(* IEC 61131-3 sources: RootPLC/crates/rootplc-stdlib/libs/Tc3_EventLogger/1.0.0, 1 file *)

(* ---- Tc3_EventLogger.st ---- *)
(* Tc3_EventLogger compatibility library for RootPLC (see library.toml).

   Written from the public library manual (TE1000 PLC Library:
   Tc3_EventLogger, version 1.6.2). RootPLC has no TwinCAT EventLogger
   service, so the blocks that talk to it are declared but not implemented
   (library.toml declare_only): calls type-check and give warning RP0120, and
   running one stops with UNSUPPORTED. FB_TcSourceInfo holds data only and is
   implemented, except ResetToDefault (it needs the instance's symbol name).

   Differences from the manual, all because the manual does not publish the
   definition:
   - interfaces used only as parameter or property types (filter
     expressions, remote logger, listener context, export settings) are
     declared without members;
   - FB_TcEventFilter has only the members the manual lists;
     FB_TcClearLoggedEventsSettings lacks SetLimit / SetSorting; the remote
     logger blocks and the ADS error conversions (E_AdsErr,
     E_HRESULTAdsErr) are left out;
   - sName of the source information is STRING(255): the manual's
     STRING(ParameterList.cSourceNameSize - 1) with the default size 256.
   TC_EVENTS is generated by TwinCAT from the project's event classes and
   is not part of this library. *)

{attribute 'qualified_only'}
TYPE TcEventSeverity : (
    Verbose  := 0,
    Info     := 1,
    Warning  := 2,
    Error    := 3,
    Critical := 4);
END_TYPE

{attribute 'qualified_only'}
TYPE TcEventConfirmationState : (
    NotSupported := 0,
    NotRequired  := 1,
    WaitForConfirmation := 2,
    Confirmed := 3,
    Reset     := 4);
END_TYPE

TYPE TcEventEntry :
STRUCT
    uuidEventClass : GUID;
    nEventId       : UDINT;
    eSeverity      : TcEventSeverity;
END_STRUCT
END_TYPE

VAR_GLOBAL CONSTANT
    EMPTY_EVENT_CLASS : GUID := (Data1 := 16#0, Data2 := 16#0, Data3 := 16#0, Data4 := [16#0, 16#0, 16#0, 16#0, 16#0, 16#0, 16#0, 16#0]);
    EMPTY_EVENT_ID    : UDINT := 16#0;
    EMPTY_SEVERITY    : TcEventSeverity := TcEventSeverity#Verbose;
    SUCCESS_EVENT     : TcEventEntry := (uuidEventClass := EMPTY_EVENT_CLASS, nEventId := EMPTY_EVENT_ID, eSeverity := EMPTY_SEVERITY);
    stLibVersion_Tc3_EventLogger : ST_LibVersion;
END_VAR

NAMESPACE GVL
VAR_GLOBAL
    nLangId_OnlineMonitoring : DINT := 1033;
END_VAR
END_NAMESPACE

NAMESPACE ParameterList
VAR_GLOBAL CONSTANT
    cSourceNameSize : UDINT(81..10000) := 256;
END_VAR
END_NAMESPACE

(* interfaces the manual names without publishing their members *)
INTERFACE I_TcRemoteEventLogger
END_INTERFACE
INTERFACE I_TcListenerContext
END_INTERFACE
INTERFACE I_TcEventFilterBase
END_INTERFACE
INTERFACE I_TcEventFilter EXTENDS I_TcEventFilterBase
END_INTERFACE
INTERFACE I_TcExpressionBase
END_INTERFACE
INTERFACE I_TcBinaryExpression
END_INTERFACE
INTERFACE I_TcLogicalExpression
END_INTERFACE
INTERFACE I_TcAlarmFilterExpression
END_INTERFACE
INTERFACE I_TcEtherCATDeviceExpression
END_INTERFACE
INTERFACE I_TcGuidCompare
END_INTERFACE
INTERFACE I_TcUDIntCompare
END_INTERFACE
INTERFACE I_TcULIntCompare
END_INTERFACE
INTERFACE I_TcJsonAttributeExpression
END_INTERFACE
INTERFACE I_TcSeverityCompare
END_INTERFACE
INTERFACE I_TcSourceInfoExpression
END_INTERFACE
INTERFACE I_TcClearLoggedEventsSettings
END_INTERFACE
INTERFACE I_TcEventExportSettings
END_INTERFACE
INTERFACE ITcEventFilterConfig
END_INTERFACE

INTERFACE I_TcSourceInfo
METHOD EqualsTo : BOOL
VAR_INPUT
    ipOther : I_TcSourceInfo;
END_VAR
END_METHOD
PROPERTY guid : GUID
GET
END_GET
END_PROPERTY
PROPERTY nId : UDINT
GET
END_GET
END_PROPERTY
PROPERTY sName : STRING(255)
GET
END_GET
END_PROPERTY
END_INTERFACE

INTERFACE I_TcArguments
METHOD AddBlob : I_TcArguments
VAR_INPUT
    pData  : PVOID;
    cbData : UINT;
END_VAR
END_METHOD
METHOD AddBool : I_TcArguments
VAR_INPUT
    value : BOOL;
END_VAR
END_METHOD
METHOD AddByte : I_TcArguments
VAR_INPUT
    value : BYTE;
END_VAR
END_METHOD
METHOD AddDINT : I_TcArguments
VAR_INPUT
    value : DINT;
END_VAR
END_METHOD
METHOD AddDWord : I_TcArguments
VAR_INPUT
    value : DWORD;
END_VAR
END_METHOD
METHOD AddEventReferenceId : I_TcArguments
VAR_INPUT
    nEventId : UDINT;
END_VAR
END_METHOD
METHOD AddEventReferenceIdGuid : I_TcArguments
VAR_INPUT
    nEventId   : UDINT;
    EventClass : GUID;
END_VAR
END_METHOD
METHOD AddINT : I_TcArguments
VAR_INPUT
    value : INT;
END_VAR
END_METHOD
METHOD AddLInt : I_TcArguments
VAR_INPUT
    value : LINT;
END_VAR
END_METHOD
METHOD AddLReal : I_TcArguments
VAR_INPUT
    value : LREAL;
END_VAR
END_METHOD
METHOD AddReal : I_TcArguments
VAR_INPUT
    value : REAL;
END_VAR
END_METHOD
METHOD AddSInt : I_TcArguments
VAR_INPUT
    value : SInt;
END_VAR
END_METHOD
METHOD AddString : I_TcArguments
VAR_IN_OUT CONSTANT
    value : STRING;
END_VAR
END_METHOD
METHOD AddUDInt : I_TcArguments
VAR_INPUT
    value : UDINT;
END_VAR
END_METHOD
METHOD AddUInt : I_TcArguments
VAR_INPUT
    value : UINT;
END_VAR
END_METHOD
METHOD AddULInt : I_TcArguments
VAR_INPUT
    value : ULINT;
END_VAR
END_METHOD
METHOD AddUSInt : I_TcArguments
VAR_INPUT
    value : USINT;
END_VAR
END_METHOD
METHOD AddWord : I_TcArguments
VAR_INPUT
    value : WORD;
END_VAR
END_METHOD
METHOD AddWString : I_TcArguments
VAR_IN_OUT CONSTANT
    value : WSTRING;
END_VAR
END_METHOD
METHOD Clear : I_TcArguments
END_METHOD
PROPERTY nCount : UDINT
GET
END_GET
END_PROPERTY
END_INTERFACE

INTERFACE I_TcEventBase
METHOD EqualsTo : BOOL
VAR_INPUT
    ipOther : I_TcEventBase;
END_VAR
END_METHOD
METHOD EqualsToEventClass : BOOL
VAR_INPUT
    OtherEventClass : GUID;
END_VAR
END_METHOD
METHOD EqualsToEventEntry : BOOL
VAR_INPUT
    OtherEventClass : GUID;
    nOtherEventID   : UDINT;
    eOtherSeverity  : TcEventSeverity;
END_VAR
END_METHOD
METHOD EqualsToEventEntryEx : BOOL
VAR_INPUT
    stOther : TcEventEntry;
END_VAR
END_METHOD
METHOD GetJsonAttribute : HRESULT
VAR_INPUT
    sJsonAttribute : REFERENCE TO STRING;
    nJsonAttribute : UDINT;
END_VAR
END_METHOD
METHOD RequestEventClassName : BOOL
VAR_INPUT
    nLangId     : DINT;
    sResult     : REFERENCE TO STRING;
    nResultSize : UDINT;
END_VAR
VAR_OUTPUT
    bError      : BOOL;
    hrErrorCode : HRESULT;
END_VAR
END_METHOD
METHOD RequestEventText : BOOL
VAR_INPUT
    nLangId     : DINT;
    sResult     : REFERENCE TO STRING;
    nResultSize : UDINT;
END_VAR
VAR_OUTPUT
    bError      : BOOL;
    hrErrorCode : HRESULT;
END_VAR
END_METHOD
PROPERTY eSeverity : TcEventSeverity
GET
END_GET
END_PROPERTY
PROPERTY EventClass : GUID
GET
END_GET
END_PROPERTY
PROPERTY ipSourceInfo : I_TcSourceInfo
GET
END_GET
END_PROPERTY
PROPERTY nEventId : UDINT
GET
END_GET
END_PROPERTY
PROPERTY stEventEntry : TcEventEntry
GET
END_GET
END_PROPERTY
END_INTERFACE

INTERFACE I_TcMessage EXTENDS I_TcEventBase
METHOD Send : HRESULT
VAR_INPUT
    nTimeStamp: ULINT;
END_VAR
END_METHOD
END_INTERFACE

INTERFACE I_Listener2
METHOD OnAlarmCleared : HRESULT
VAR_INPUT
    fbEvent : REFERENCE TO FB_TcEvent;
END_VAR
END_METHOD
METHOD OnAlarmConfirmed : HRESULT
VAR_INPUT
    fbEvent : REFERENCE TO FB_TcEvent;
END_VAR
END_METHOD
METHOD OnAlarmDisposed : HRESULT
VAR_INPUT
    fbEvent : REFERENCE TO FB_TcEvent;
END_VAR
END_METHOD
METHOD OnAlarmRaised : HRESULT
VAR_INPUT
    fbEvent : REFERENCE TO FB_TcEvent;
END_VAR
END_METHOD
METHOD OnMessageSent : HRESULT
VAR_INPUT
    fbEvent : REFERENCE TO FB_TcEvent;
END_VAR
END_METHOD
END_INTERFACE

FUNCTION_BLOCK FB_AsyncStrResult
METHOD GetString : BOOL
VAR_INPUT
    sResult : REFERENCE TO STRING;
    nResult : UDINT;
END_VAR
END_METHOD
PROPERTY bBusy : BOOL
GET
END_GET
END_PROPERTY
PROPERTY bError : BOOL
GET
END_GET
END_PROPERTY
PROPERTY hrErrorCode : HRESULT
GET
END_GET
END_PROPERTY
END_FUNCTION_BLOCK

FUNCTION_BLOCK FB_TcCauseRemedy
METHOD GetCause : BOOL
VAR_INPUT
    sResult     : REFERENCE TO STRING;
    nResult     : UDINT; (* buffer size in bytes *)
END_VAR
END_METHOD
METHOD GetId : BOOL
VAR_INPUT
    sResult  : REFERENCE TO STRING;
    nResult  : UDINT; (* buffer size in bytes *)
END_VAR
END_METHOD
METHOD GetRemedy : BOOL
VAR_INPUT
    sResult      : REFERENCE TO STRING;
    nResult      : UDINT; (* buffer size in bytes *)
END_VAR
END_METHOD
METHOD Release : HRESULT
END_METHOD
END_FUNCTION_BLOCK

FUNCTION_BLOCK FB_TcDetail
METHOD Release : HRESULT
END_METHOD
METHOD GetComment : BOOL
VAR_INPUT
    sResult       : REFERENCE TO STRING;
    nResult       : UDINT; (* buffer size in bytes *)
END_VAR
END_METHOD
METHOD GetName : BOOL
VAR_INPUT
    sResult    : REFERENCE TO STRING;
    nResult    : UDINT; (* buffer size in bytes *)
END_VAR
END_METHOD
METHOD GetText : BOOL
VAR_INPUT
    sResult    : REFERENCE TO STRING;
    nResult    : UDINT; (* buffer size in bytes *)
END_VAR
END_METHOD
END_FUNCTION_BLOCK

FUNCTION_BLOCK FB_RequestCauseRemedy
METHOD Clear
END_METHOD
METHOD Get        : HRESULT
VAR_INPUT
    nIndex        : UDINT;
    fbCauseRemedy : REFERENCE TO FB_TcCauseRemedy;
END_VAR
END_METHOD
METHOD Request : HRESULT
VAR_INPUT
    eventClass : GUID;
    nEventId   : UDINT;
    nLangId    : DINT; (* English(US)=1033 ; German(Germay)=1031 *)
END_VAR
END_METHOD
METHOD RequestRemote : HRESULT
VAR_INPUT
    ipRemoteLogger   : I_TcRemoteEventLogger;
    eventClass       : GUID;
    nEventId         : UDINT;
    nLangId          : DINT; (* English(US)=1033 ; German(Germay)=1031 *)
END_VAR
END_METHOD
PROPERTY bBusy : BOOL
GET
END_GET
END_PROPERTY
PROPERTY bError : BOOL
GET
END_GET
END_PROPERTY
PROPERTY hrErrorCode : HRESULT
GET
END_GET
END_PROPERTY
PROPERTY nCount : UDINT
GET
END_GET
END_PROPERTY
END_FUNCTION_BLOCK

FUNCTION_BLOCK FB_RequestEventClassDetails
METHOD Clear
END_METHOD
METHOD Get   : HRESULT
VAR_INPUT
    nIndex   : UDINT;
    fbDetail : REFERENCE TO FB_TcDetail;
END_VAR
END_METHOD
METHOD Request : HRESULT
VAR_INPUT
    eventClass : GUID;
    nLangId    : DINT; (* English(US)=1033 ; German(Germay)=1031 *)
END_VAR
END_METHOD
METHOD RequestRemote : HRESULT
VAR_INPUT
    ipRemoteLogger   : I_TcRemoteEventLogger;
    eventClass       : GUID;
    nLangId          : DINT; (* English(US)=1033 ; German(Germay)=1031 *)
END_VAR
END_METHOD
PROPERTY bBusy : BOOL
GET
END_GET
END_PROPERTY
PROPERTY bError : BOOL
GET
END_GET
END_PROPERTY
PROPERTY hrErrorCode : HRESULT
GET
END_GET
END_PROPERTY
PROPERTY nCount : UDINT
GET
END_GET
END_PROPERTY
END_FUNCTION_BLOCK

FUNCTION_BLOCK FB_RequestEventClassName
METHOD Clear
END_METHOD
METHOD GetString : BOOL
VAR_INPUT
    sResult : REFERENCE TO STRING;
    nResult : UDINT;
END_VAR
END_METHOD
METHOD Request : HRESULT
VAR_INPUT
    eventClass : GUID;
    nLangId    : DINT;
END_VAR
END_METHOD
METHOD RequestRemote : HRESULT
VAR_INPUT
    ipRemoteLogger   : I_TcRemoteEventLogger;
    eventClass       : GUID;
    nLangId          : DINT; (* English(US)=1033 ; German(Germay)=1031 *)
END_VAR
END_METHOD
PROPERTY bBusy : BOOL
GET
END_GET
END_PROPERTY
PROPERTY bError : BOOL
GET
END_GET
END_PROPERTY
PROPERTY hrErrorCode : HRESULT
GET
END_GET
END_PROPERTY
END_FUNCTION_BLOCK

FUNCTION_BLOCK FB_RequestEventDetails
METHOD Clear
END_METHOD
METHOD Get   : HRESULT
VAR_INPUT
    nIndex   : UDINT;
    fbDetail : REFERENCE TO FB_TcDetail;
END_VAR
END_METHOD
METHOD Request : HRESULT
VAR_INPUT
    eventClass : GUID;
    nEventId   : UDINT;
    nLangId    : DINT; (* English(US)=1033 ; German(Germay)=1031 *)
END_VAR
END_METHOD
METHOD RequestRemote : HRESULT
VAR_INPUT
    ipRemoteLogger   : I_TcRemoteEventLogger;
    eventClass       : GUID;
    nEventId         : UDINT;
    nLangId          : DINT; (* English(US)=1033 ; German(Germay)=1031 *)
END_VAR
END_METHOD
PROPERTY bBusy : BOOL
GET
END_GET
END_PROPERTY
PROPERTY bError : BOOL
GET
END_GET
END_PROPERTY
PROPERTY hrErrorCode : HRESULT
GET
END_GET
END_PROPERTY
PROPERTY nCount : UDINT
GET
END_GET
END_PROPERTY
END_FUNCTION_BLOCK

FUNCTION_BLOCK FB_RequestEventText
METHOD GetString : BOOL
VAR_INPUT
    sResult : REFERENCE TO STRING;
    nResult : UDINT;
END_VAR
END_METHOD
METHOD Request : BOOL
VAR_INPUT
    eventClass : GUID;
    nEventId   : UDINT;
    nLangId    : DINT;
    ipArgs     : I_TcArguments;
END_VAR
END_METHOD
METHOD RequestRemote : HRESULT
VAR_INPUT
    ipRemoteLogger   : I_TcRemoteEventLogger;
    eventClass       : GUID;
    nEventId         : UDINT;
    nLangId          : DINT;
    ipArgs           : I_TcArguments;
END_VAR
END_METHOD
METHOD Clear
END_METHOD
PROPERTY bBusy : BOOL
GET
END_GET
END_PROPERTY
PROPERTY bError : BOOL
GET
END_GET
END_PROPERTY
PROPERTY hrErrorCode : HRESULT
GET
END_GET
END_PROPERTY
END_FUNCTION_BLOCK

FUNCTION_BLOCK FB_RequestTranslation
METHOD GetString : BOOL
VAR_INPUT
    sResult : REFERENCE TO STRING;
    nResult : UDINT;
END_VAR
END_METHOD
METHOD Request : BOOL
VAR_INPUT
    eventClass : GUID;
END_VAR
VAR_IN_OUT CONSTANT
    text       : STRING;
END_VAR
VAR_INPUT
    nLangId    : DINT;
    ipArgs     : I_TcArguments;
END_VAR
END_METHOD
METHOD RequestRemote : HRESULT
VAR_INPUT
    ipRemoteLogger   : I_TcRemoteEventLogger;
    eventClass       : GUID;
END_VAR
VAR_IN_OUT CONSTANT
    text             : STRING;
END_VAR
VAR_INPUT
    nLangId          : DINT;
    ipArgs           : I_TcArguments;
END_VAR
END_METHOD
METHOD Clear
END_METHOD
PROPERTY bBusy : BOOL
GET
END_GET
END_PROPERTY
PROPERTY bError : BOOL
GET
END_GET
END_PROPERTY
PROPERTY hrErrorCode : HRESULT
GET
END_GET
END_PROPERTY
END_FUNCTION_BLOCK

FUNCTION_BLOCK FB_TcEventBase
METHOD EqualsTo : BOOL
VAR_INPUT
    ipOther : I_TcEventBase;
END_VAR
END_METHOD
METHOD EqualsToEventClass : BOOL
VAR_INPUT
    OtherEventClass : GUID;
END_VAR
END_METHOD
METHOD EqualsToEventEntry : BOOL
VAR_INPUT
    OtherEventClass : GUID;
    nOtherEventID   : UDINT;
    eOtherSeverity  : TcEventSeverity;
END_VAR
END_METHOD
METHOD EqualsToEventEntryEx : BOOL
VAR_INPUT
    stOther : TcEventEntry;
END_VAR
END_METHOD
METHOD GetJsonAttribute : HRESULT
VAR_INPUT
    sJsonAttribute : REFERENCE TO STRING;
    nJsonAttribute : UDINT;
END_VAR
END_METHOD
METHOD Release : HRESULT
END_METHOD
METHOD RequestEventClassName : BOOL
VAR_INPUT
    nLangId     : DINT;
    sResult     : REFERENCE TO STRING;
    nResultSize : UDINT;
END_VAR
VAR_OUTPUT
    bError      : BOOL;
    hrErrorCode : HRESULT;
END_VAR
END_METHOD
METHOD RequestEventText : BOOL
VAR_INPUT
    nLangId     : DINT;
    sResult     : REFERENCE TO STRING;
    nResultSize : UDINT;
END_VAR
VAR_OUTPUT
    bError      : BOOL;
    hrErrorCode : HRESULT;
END_VAR
END_METHOD
PROPERTY eSeverity : TcEventSeverity
GET
END_GET
END_PROPERTY
PROPERTY EventClass : GUID
GET
END_GET
END_PROPERTY
PROPERTY ipArguments : I_TcArguments
GET
END_GET
END_PROPERTY
PROPERTY ipSourceInfo : I_TcSourceInfo
GET
END_GET
END_PROPERTY
PROPERTY nEventId : UDINT
GET
END_GET
END_PROPERTY
PROPERTY nUniqueId : UDINT
GET
END_GET
END_PROPERTY
PROPERTY stEventEntry : TcEventEntry
GET
END_GET
END_PROPERTY
END_FUNCTION_BLOCK

FUNCTION_BLOCK FB_TcEvent EXTENDS FB_TcEventBase IMPLEMENTS I_TcEventBase
PROPERTY nTimestamp : ULINT
GET
END_GET
END_PROPERTY
END_FUNCTION_BLOCK

FUNCTION_BLOCK FB_TcMessage EXTENDS FB_TcEventBase IMPLEMENTS I_TcMessage
METHOD Create : HRESULT
VAR_INPUT
    eventClass   : GUID;
    nEventId     : UDINT;
    eSeverity    : TcEventSeverity;
    ipSourceInfo : I_TcSourceInfo := 0;
END_VAR
END_METHOD
METHOD CreateEx : HRESULT
VAR_INPUT
    stEventEntry : TcEventEntry;
    ipSourceInfo : I_TcSourceInfo := 0;
END_VAR
END_METHOD
METHOD SetJsonAttribute : HRESULT
VAR_IN_OUT CONSTANT
    sJsonAttribute : STRING;
END_VAR
END_METHOD
METHOD Send : HRESULT
VAR_INPUT
    nTimeStamp: ULINT;
END_VAR
END_METHOD
PROPERTY nTimeSent : ULINT
GET
END_GET
END_PROPERTY
END_FUNCTION_BLOCK

FUNCTION_BLOCK FB_TcAlarm EXTENDS FB_TcEventBase
METHOD Clear : HRESULT
VAR_INPUT
    nTimeStamp         : ULINT;
    bResetConfirmation : BOOL;
END_VAR
END_METHOD
METHOD Confirm : HRESULT
VAR_INPUT
    nTimeStamp: ULINT;
END_VAR
END_METHOD
METHOD Create : HRESULT
VAR_INPUT
    eventClass        : GUID;
    nEventId          : UDINT;
    eSeverity         : TcEventSeverity;
    bWithConfirmation : BOOL;
    ipSourceInfo      : I_TcSourceInfo;
END_VAR
END_METHOD
METHOD CreateEx : HRESULT
VAR_INPUT
    stEventEntry      : TcEventEntry;
    bWithConfirmation : BOOL;
    ipSourceInfo      : I_TcSourceInfo;
END_VAR
END_METHOD
METHOD Raise : HRESULT
VAR_INPUT
    nTimeStamp : ULINT;
END_VAR
END_METHOD
METHOD SetJsonAttribute : HRESULT
VAR_IN_OUT CONSTANT
    sJsonAttribute : STRING;
END_VAR
END_METHOD
PROPERTY bRaised : BOOL
GET
END_GET
END_PROPERTY
PROPERTY bActive : BOOL
GET
END_GET
END_PROPERTY
PROPERTY eConfirmationState : TcEventConfirmationState
GET
END_GET
END_PROPERTY
PROPERTY nTimeCleared : ULINT
GET
END_GET
END_PROPERTY
PROPERTY nTimeConfirmed : ULINT
GET
END_GET
END_PROPERTY
PROPERTY nTimeRaised : ULINT
GET
END_GET
END_PROPERTY
END_FUNCTION_BLOCK

FUNCTION_BLOCK FB_TcArguments IMPLEMENTS I_TcArguments
METHOD IsEmpty : BOOL
END_METHOD
METHOD AddBlob : I_TcArguments
VAR_INPUT
    pData  : PVOID;
    cbData : UINT;
END_VAR
END_METHOD
METHOD AddBool : I_TcArguments
VAR_INPUT
    value : BOOL;
END_VAR
END_METHOD
METHOD AddByte : I_TcArguments
VAR_INPUT
    value : BYTE;
END_VAR
END_METHOD
METHOD AddDINT : I_TcArguments
VAR_INPUT
    value : DINT;
END_VAR
END_METHOD
METHOD AddDWord : I_TcArguments
VAR_INPUT
    value : DWORD;
END_VAR
END_METHOD
METHOD AddEventReferenceId : I_TcArguments
VAR_INPUT
    nEventId : UDINT;
END_VAR
END_METHOD
METHOD AddEventReferenceIdGuid : I_TcArguments
VAR_INPUT
    nEventId   : UDINT;
    EventClass : GUID;
END_VAR
END_METHOD
METHOD AddINT : I_TcArguments
VAR_INPUT
    value : INT;
END_VAR
END_METHOD
METHOD AddLInt : I_TcArguments
VAR_INPUT
    value : LINT;
END_VAR
END_METHOD
METHOD AddLReal : I_TcArguments
VAR_INPUT
    value : LREAL;
END_VAR
END_METHOD
METHOD AddReal : I_TcArguments
VAR_INPUT
    value : REAL;
END_VAR
END_METHOD
METHOD AddSInt : I_TcArguments
VAR_INPUT
    value : SInt;
END_VAR
END_METHOD
METHOD AddString : I_TcArguments
VAR_IN_OUT CONSTANT
    value : STRING;
END_VAR
END_METHOD
METHOD AddUDInt : I_TcArguments
VAR_INPUT
    value : UDINT;
END_VAR
END_METHOD
METHOD AddUInt : I_TcArguments
VAR_INPUT
    value : UINT;
END_VAR
END_METHOD
METHOD AddULInt : I_TcArguments
VAR_INPUT
    value : ULINT;
END_VAR
END_METHOD
METHOD AddUSInt : I_TcArguments
VAR_INPUT
    value : USINT;
END_VAR
END_METHOD
METHOD AddWord : I_TcArguments
VAR_INPUT
    value : WORD;
END_VAR
END_METHOD
METHOD AddWString : I_TcArguments
VAR_IN_OUT CONSTANT
    value : WSTRING;
END_VAR
END_METHOD
METHOD Clear : I_TcArguments
END_METHOD
PROPERTY nCount : UDINT
GET
END_GET
END_PROPERTY
END_FUNCTION_BLOCK

FUNCTION_BLOCK FB_TcEventLogger
METHOD ClearAlarms     : HRESULT
VAR_INPUT
    nTimeStamp         : ULINT := 0;
    bResetConfirmation : BOOL  := FALSE;
    ipFilter           : I_TcEventFilter;
END_VAR
END_METHOD
METHOD ClearAllAlarms : HRESULT
VAR_INPUT
    nTimeStamp         : ULINT := 0;
    bResetConfirmation : BOOL := FALSE;
END_VAR
END_METHOD
METHOD ClearLoggedEvents : BOOL
VAR_INPUT
    ipClearSettings      : I_TcClearLoggedEventsSettings;
END_VAR
VAR_OUTPUT
    bError               : BOOL;
    hrErrorCode          : HRESULT;
END_VAR
END_METHOD
METHOD ConfirmAlarms : HRESULT
VAR_INPUT
    nTimeStamp       : ULINT := 0;
    ipFilter         : I_TcEventFilter;
END_VAR
END_METHOD
METHOD ConfirmAllAlarms : HRESULT
VAR_INPUT
    nTimeStamp : ULINT := 0;
END_VAR
END_METHOD
METHOD ExportLoggedEvents : BOOL
VAR_IN_OUT CONSTANT
    sFileName             : STRING;
END_VAR
VAR_INPUT
ipExportSettings          : I_TcEventExportSettings;
END_VAR
VAR_OUTPUT
    bError                : BOOL;
    hrErrorCode           : HRESULT;
END_VAR
END_METHOD
METHOD GetAlarm : HRESULT
VAR_INPUT
    eventClass   : GUID;
    nEventId     : UDINT;
    ipSourceInfo : I_TcSourceInfo := 0;
    fbAlarm      : REFERENCE TO FB_TcAlarm;
END_VAR
END_METHOD
METHOD GetAlarmEx : HRESULT
VAR_INPUT
    stEventEntry : TcEventEntry;
    ipSourceInfo : I_TcSourceInfo := 0; (* optional *)
    fbAlarm      : REFERENCE TO FB_TcAlarm;
END_VAR
END_METHOD
METHOD IsAlarmRaised : BOOL
VAR_INPUT
    eventClass   : GUID;
    nEventId     : UDINT;
    ipSourceInfo : I_TcSourceInfo := 0;
END_VAR
END_METHOD
METHOD IsAlarmRaisedEx : BOOL
VAR_INPUT
    stEventEntry : TcEventEntry;
    ipSourceInfo : I_TcSourceInfo := 0;
END_VAR
END_METHOD
METHOD SendMessage : HRESULT
VAR_INPUT
    eventClass    : GUID;
    nEventId      : UDINT;
    eSeverity     : TcEventSeverity;
    ipSourceInfo  : I_TcSourceInfo := 0;
    nTimeStamp    : ULINT := 0;
    ipArguments   : I_TcArguments := 0;
END_VAR
END_METHOD
METHOD SendMessage2 : HRESULT
VAR_INPUT
    eventClass      : GUID;
    nEventId        : UDINT;
    eSeverity       : TcEventSeverity;
    ipSourceInfo    : I_TcSourceInfo := 0;
    nTimeStamp      : ULINT := 0;
    ipArguments     : I_TcArguments := 0;
END_VAR
VAR_IN_OUT CONSTANT
    sJsonAttribute  : STRING;
END_VAR
END_METHOD
METHOD SendMessageEx : HRESULT
VAR_INPUT
    stEventEntry : TcEventEntry;
    ipSourceInfo : I_TcSourceInfo := 0;
    nTimeStamp   : ULINT := 0;
    ipArguments  : I_TcArguments := 0;
END_VAR
END_METHOD
METHOD SendMessageEx2 : HRESULT
VAR_INPUT
    stEventEntry      : TcEventEntry;
    ipSourceInfo      : I_TcSourceInfo := 0;
    nTimeStamp        : ULINT := 0;
    ipArguments       : I_TcArguments := 0;
END_VAR
VAR_IN_OUT CONSTANT
    sJsonAttribute    : STRING;
END_VAR
END_METHOD
END_FUNCTION_BLOCK

FUNCTION_BLOCK FB_ListenerBase2 IMPLEMENTS I_Listener2
METHOD Execute : HRESULT
END_METHOD
METHOD OnAlarmCleared : HRESULT
VAR_INPUT
    fbEvent : REFERENCE TO FB_TcEvent;
END_VAR
END_METHOD
METHOD OnAlarmConfirmed : HRESULT
VAR_INPUT
    fbEvent : REFERENCE TO FB_TcEvent;
END_VAR
END_METHOD
METHOD OnAlarmDisposed : HRESULT
VAR_INPUT
    fbEvent : REFERENCE TO FB_TcEvent;
END_VAR
END_METHOD
METHOD OnAlarmRaised : HRESULT
VAR_INPUT
    fbEvent : REFERENCE TO FB_TcEvent;
END_VAR
END_METHOD
METHOD OnMessageSent : HRESULT
VAR_INPUT
    fbEvent : REFERENCE TO FB_TcEvent;
END_VAR
END_METHOD
METHOD Subscribe : HRESULT
VAR_INPUT
    ipMessageFilterConfig : POINTER TO ITcEventFilterConfig;
    ipAlarmFilterConfig   : POINTER TO ITcEventFilterConfig;
END_VAR
END_METHOD
METHOD Subscribe2 : HRESULT
VAR_INPUT
    ipEventFilter : I_TcEventFilterBase;
END_VAR
END_METHOD
METHOD Unsubscribe : HRESULT
END_METHOD
END_FUNCTION_BLOCK

FUNCTION F_GetEventClassName : HRESULT
VAR_INPUT
    nLangId     : DINT;
    fbEventBase : REFERENCE TO FB_TcEventBase;
END_VAR
VAR_IN_OUT
    fbResult : FB_AsyncStrResult;
END_VAR
END_FUNCTION

FUNCTION F_GetEventText : HRESULT
VAR_INPUT
    nLangId     : DINT;
    fbEventBase : REFERENCE TO FB_TcEventBase;
END_VAR
VAR_IN_OUT
    fbResult : FB_AsyncStrResult;
END_VAR
END_FUNCTION

FUNCTION_BLOCK FB_TcSourceInfo IMPLEMENTS I_TcSourceInfo
VAR
    _guid  : GUID;
    _nId   : UDINT;
    _sName : STRING(255);
END_VAR
METHOD Clear
VAR
    empty : GUID;
END_VAR
_guid := empty;
_nId := 0;
_sName := '';
END_METHOD
METHOD ExtendName : BOOL
VAR_INPUT
    sExtension : STRING(255);
END_VAR
ExtendName := LEN(_sName) + LEN(sExtension) <= 255;
_sName := CONCAT(_sName, sExtension);
END_METHOD
METHOD ResetToDefault
END_METHOD
METHOD EqualsTo : BOOL
VAR_INPUT
    ipOther : I_TcSourceInfo;
END_VAR
VAR
    g : GUID;
    i : INT;
END_VAR
IF ipOther = 0 THEN
    RETURN;
END_IF
g := ipOther.guid;
EqualsTo := g.Data1 = _guid.Data1 AND g.Data2 = _guid.Data2 AND g.Data3 = _guid.Data3
    AND ipOther.nId = _nId AND ipOther.sName = _sName;
FOR i := 0 TO 7 DO
    EqualsTo := EqualsTo AND g.Data4[i] = _guid.Data4[i];
END_FOR
END_METHOD
PROPERTY guid : GUID
GET
    guid := _guid;
END_GET
SET
    _guid := guid;
END_SET
END_PROPERTY
PROPERTY nId : UDINT
GET
    nId := _nId;
END_GET
SET
    _nId := nId;
END_SET
END_PROPERTY
PROPERTY sName : STRING(255)
GET
    sName := _sName;
END_GET
SET
    _sName := sName;
END_SET
END_PROPERTY
END_FUNCTION_BLOCK

FUNCTION_BLOCK FB_TcEventFilter IMPLEMENTS I_TcEventFilter, I_TcExpressionBase
METHOD Clear : I_TcBinaryExpression
END_METHOD
METHOD FilterExpression : I_TcLogicalExpression
VAR_INPUT
    ipExpression : I_TcEventFilterBase;
END_VAR
END_METHOD
METHOD IsAlarm : I_TcLogicalExpression
END_METHOD
METHOD IsMessage : I_TcLogicalExpression
END_METHOD
METHOD NOT_OP : I_TcBinaryExpression
END_METHOD
PROPERTY AlarmState : I_TcAlarmFilterExpression
GET
END_GET
END_PROPERTY
PROPERTY EtherCATDevice : I_TcEtherCATDeviceExpression
GET
END_GET
END_PROPERTY
PROPERTY EventClass : I_TcGuidCompare
GET
END_GET
END_PROPERTY
PROPERTY EventId : I_TcUDIntCompare
GET
END_GET
END_PROPERTY
PROPERTY JsonAttribute : I_TcJsonAttributeExpression
GET
END_GET
END_PROPERTY
PROPERTY Severity : I_TcSeverityCompare
GET
END_GET
END_PROPERTY
PROPERTY Source : I_TcSourceInfoExpression
GET
END_GET
END_PROPERTY
PROPERTY TimeCleared : I_TcULIntCompare
GET
END_GET
END_PROPERTY
PROPERTY TimeConfirmed : I_TcULIntCompare
GET
END_GET
END_PROPERTY
PROPERTY TimeRaised : I_TcULIntCompare
GET
END_GET
END_PROPERTY
END_FUNCTION_BLOCK

FUNCTION_BLOCK FB_TcClearLoggedEventsSettings IMPLEMENTS I_TcClearLoggedEventsSettings
METHOD AddFilter : HRESULT
VAR_INPUT
    ipEventFilter : I_TcEventFilter;
END_VAR
END_METHOD
METHOD Clear : HRESULT
END_METHOD
END_FUNCTION_BLOCK
